(* IEC 61131-3 sources: codesys-to-s7/tests/corpus/C2S7-TYPE-DATE/pos, 1 file *)

(* ---- input.st ---- *)
FUNCTION_BLOCK FB_Case
VAR
    w : WORD;
    dtNow : DT;
END_VAR
w := DWORD_TO_WORD(DT_TO_DWORD(dtNow));
END_FUNCTION_BLOCK
